(*!
<summary>Selects one independently reported scenario in the WorkflowComprehensiveTest group.</summary>
*)
{attribute 'qualified_only'}
{attribute 'strict'}
TYPE WORKFLOW_COMPREHENSIVE_TEST_SCENARIO :
(
	END_TO_END_COMPREHENSIVE_SCENARIO,
	WORKFLOW_RESET,
	WORKFLOW_CANCEL,
	PARALLEL_ACTIVITY_WAIT_ALL,
	PARALLEL_ACTIVITY_WAIT_ANY,
	NOT_CONDITION,
	COMPARE_VARIABLE_CONDITION,
	MIXED_NUMERIC_COMPARISON,
	MIXED_TEXT_COMPARISON,
	STANDARD_COMPARISON_FALLBACK,
	INCOMPATIBLE_COMPARISON_PAIRS,
	DIRECT_WORKFLOW_DYNAMIC_CREATION,
	ACTIVITY_VARIABLE_SCOPING_AND_SHADOWING,
	VARIABLE_REGISTRATION_VALIDATION
);
END_TYPE

(* stored: Version 1.1.0.1
   DUT WORKFLOW_COMPREHENSIVE_TEST_SCENARIO: Id {7d2c1bf6-47d2-4d1e-9658-01c5c1d32597} *)
